(* IEC 61131-3 sources: RoboFlex-Cell/plc/codesys, 6 files *)

(* ---- FB_Alarm.st ---- *)
FUNCTION_BLOCK FB_Alarm
VAR_INPUT
    Trip : BOOL;
    Code : UINT;
    ResetAccepted : BOOL;
END_VAR
VAR_OUTPUT
    Active : BOOL;
    LatchedCode : UINT;
END_VAR
IF Trip THEN
    IF NOT Active THEN
        LatchedCode := Code;
    END_IF;
    Active := TRUE;
ELSIF ResetAccepted THEN
    Active := FALSE;
    LatchedCode := 0;
END_IF;
END_FUNCTION_BLOCK

(* ---- FB_Conveyor.st ---- *)
FUNCTION_BLOCK FB_Conveyor
VAR_INPUT
    RunRequest : BOOL;
    SafeEnable : BOOL;
    JamDetected : BOOL;
END_VAR
VAR_OUTPUT
    MotorRun : BOOL;
END_VAR
MotorRun := RunRequest AND SafeEnable AND NOT JamDetected;
END_FUNCTION_BLOCK

(* ---- FB_Gripper.st ---- *)
FUNCTION_BLOCK FB_Gripper
VAR_INPUT
    CloseRequest : BOOL;
    ClosedFeedback : BOOL;
    OpenFeedback : BOOL;
    SafeEnable : BOOL;
    Reset : BOOL;
END_VAR
VAR_OUTPUT
    CloseValve : BOOL;
    AtPosition : BOOL;
    Error : BOOL;
END_VAR
VAR
    FeedbackTimer : TON;
END_VAR
(* Hold the last valve command on a software safety stop; never drop a part.
   A physical safety circuit requires an independently assessed pneumatic design. *)
IF SafeEnable THEN
    CloseValve := CloseRequest;
END_IF;
AtPosition := (CloseRequest AND ClosedFeedback) OR (NOT CloseRequest AND OpenFeedback);
FeedbackTimer(IN := SafeEnable AND NOT AtPosition, PT := T#500ms);
IF Reset THEN
    Error := FALSE;
ELSIF FeedbackTimer.Q THEN
    Error := TRUE;
END_IF;
END_FUNCTION_BLOCK

(* ---- FB_Robot.st ---- *)
FUNCTION_BLOCK FB_Robot
VAR_INPUT
    Execute : BOOL;
    SafeEnable : BOOL;
    Reset : BOOL;
    Ready : BOOL;
    Running : BOOL;
    Complete : BOOL;
    RobotError : BOOL;
END_VAR
VAR_OUTPUT
    Start : BOOL;
    Ack : BOOL;
    Stop : BOOL;
    Done : BOOL;
    Error : BOOL;
    ErrorId : UINT;
END_VAR
VAR
    Phase : UINT;
    StartEdge : R_TRIG;
    StartTimer : TON;
    MotionTimer : TON;
    AckTimer : TON;
END_VAR

StartEdge(CLK := Execute);
StartTimer(IN := Phase = 10, PT := T#500ms);
MotionTimer(IN := Phase = 20, PT := T#6s);
AckTimer(IN := Phase = 30, PT := T#500ms);
Start := FALSE;
Ack := FALSE;
Stop := NOT SafeEnable;

IF Reset AND SafeEnable THEN
    Phase := 0;
    Done := FALSE;
    Error := FALSE;
    ErrorId := 0;
ELSIF NOT SafeEnable THEN
    Phase := 0;
    Done := FALSE;
ELSIF RobotError THEN
    Error := TRUE;
    ErrorId := 3;
END_IF;

IF SafeEnable AND NOT Reset AND NOT Error THEN
    CASE Phase OF
        0:
            IF StartEdge.Q THEN
                IF Ready AND NOT Complete AND NOT Running THEN
                    Phase := 10;
                ELSE
                    Error := TRUE;
                    ErrorId := 3;
                END_IF;
            END_IF;
        10:
            Start := TRUE;
            IF Running THEN
                Start := FALSE;
                Phase := 20;
            ELSIF StartTimer.Q THEN
                Error := TRUE;
                ErrorId := 4;
            END_IF;
        20:
            IF Complete AND NOT Running THEN
                Phase := 30;
            ELSIF MotionTimer.Q THEN
                Error := TRUE;
                ErrorId := 4;
            END_IF;
        30:
            Ack := TRUE;
            IF NOT Complete AND Ready THEN
                Ack := FALSE;
                Done := TRUE;
                Phase := 40;
            ELSIF AckTimer.Q THEN
                Error := TRUE;
                ErrorId := 4;
            END_IF;
        40:
            IF NOT Execute THEN
                Done := FALSE;
                Phase := 0;
            END_IF;
    END_CASE;
END_IF;
IF Error THEN
    Start := FALSE;
    Ack := FALSE;
    Stop := TRUE;
END_IF;
END_FUNCTION_BLOCK

(* ---- FB_Sequence.st ---- *)
FUNCTION_BLOCK FB_Sequence
VAR_INPUT
    StartButton : BOOL;
    StopButton : BOOL;
    ResetButton : BOOL;
    ManualPartClear : BOOL;
    SafetyOK : BOOL;
    HeartbeatOK : BOOL;
    PartDetected : BOOL;
    JamDetected : BOOL;
    VisionDone : BOOL;
    VisionError : BOOL;
    VisionErrorId : UINT;
    RobotDone : BOOL;
    RobotError : BOOL;
    RobotErrorId : UINT;
    GripperClosed : BOOL;
    GripperOpen : BOOL;
    GripperError : BOOL;
    QualityOK : BOOL;
END_VAR
VAR_OUTPUT
    State : UINT; (* 0 idle, 30 wait, 40 vision, 50 pick, 55 grip, 60 place,
                     65 release, 70 check, 75 home, 80 complete, 900 error *)
    ConveyorRequest : BOOL;
    VisionExecute : BOOL;
    RobotExecute : BOOL;
    JobNumber : UINT; (* 1 pick, 2 place, 3 home; pose data sent separately *)
    CloseRequest : BOOL;
    AlarmCode : UINT;
    ResetAccepted : BOOL;
    OKCount : UDINT;
    NGCount : UDINT;
END_VAR
VAR
    StartEdge : R_TRIG;
    ResetEdge : R_TRIG;
    StateTimer : TON;
    LastState : UINT;
    TripCode : UINT;
END_VAR

StartEdge(CLK := StartButton);
ResetEdge(CLK := ResetButton);
StateTimer(IN := State = LastState AND State <> 0 AND State <> 900, PT := T#2s);
LastState := State;
ResetAccepted := FALSE;
TripCode := 0;
ConveyorRequest := FALSE;
VisionExecute := FALSE;
RobotExecute := FALSE;

IF NOT SafetyOK THEN
    TripCode := 10; (* actual E-stop/door distinction belongs in mapped safety status *)
ELSIF State <> 0 AND State <> 900 THEN
    IF NOT HeartbeatOK THEN TripCode := 7;
    ELSIF StopButton THEN TripCode := 13;
    ELSIF RobotError THEN TripCode := RobotErrorId;
    ELSIF VisionError THEN TripCode := VisionErrorId;
    ELSIF GripperError THEN TripCode := 5;
    ELSIF JamDetected THEN TripCode := 9;
    END_IF;
END_IF;

IF TripCode <> 0 AND State <> 900 THEN
    AlarmCode := TripCode;
    State := 900;
END_IF;

CASE State OF
    0:
        IF StartEdge.Q AND SafetyOK AND HeartbeatOK AND NOT JamDetected THEN State := 30; END_IF;
    30:
        ConveyorRequest := TRUE;
        IF PartDetected THEN
            ConveyorRequest := FALSE;
            State := 40;
        ELSIF StateTimer.Q THEN
            AlarmCode := 8;
            State := 900;
        END_IF;
    40:
        VisionExecute := TRUE;
        IF VisionDone THEN State := 50; END_IF;
    50:
        JobNumber := 1;
        RobotExecute := TRUE;
        IF RobotDone THEN State := 55; END_IF;
    55:
        CloseRequest := TRUE;
        IF GripperClosed THEN State := 60; END_IF;
    60:
        JobNumber := 2;
        RobotExecute := TRUE;
        IF RobotDone THEN State := 65; END_IF;
    65:
        CloseRequest := FALSE;
        IF GripperOpen THEN State := 70; END_IF;
    70:
        IF QualityOK THEN State := 75;
        ELSIF StateTimer.Q THEN
            NGCount := NGCount + 1;
            AlarmCode := 6;
            State := 900;
        END_IF;
    75:
        JobNumber := 3;
        RobotExecute := TRUE;
        IF RobotDone THEN State := 80; END_IF;
    80:
        OKCount := OKCount + 1;
        State := 30;
    900:
        IF ResetEdge.Q AND SafetyOK AND HeartbeatOK AND NOT JamDetected AND ManualPartClear THEN
            ResetAccepted := TRUE;
            CloseRequest := FALSE;
            AlarmCode := 0;
            State := 0;
        END_IF;
END_CASE;
IF State = 900 THEN
    ConveyorRequest := FALSE;
    VisionExecute := FALSE;
    RobotExecute := FALSE;
END_IF;
END_FUNCTION_BLOCK

(* ---- FB_Vision.st ---- *)
FUNCTION_BLOCK FB_Vision
VAR_INPUT
    Execute : BOOL;
    SafeEnable : BOOL;
    Connected : BOOL;
    ResultValid : BOOL;
    ResultOK : BOOL;
    Reset : BOOL;
END_VAR
VAR_OUTPUT
    Trigger : BOOL;
    Ack : BOOL;
    Done : BOOL;
    Error : BOOL;
    ErrorId : UINT;
END_VAR
VAR
    Phase : UINT;
    Edge : R_TRIG;
    ResultTimer : TON;
    ClearTimer : TON;
END_VAR
Edge(CLK := Execute);
ResultTimer(IN := Phase = 10, PT := T#1s);
ClearTimer(IN := Phase = 20, PT := T#500ms);
Trigger := FALSE;
Ack := FALSE;
IF Reset OR NOT SafeEnable THEN
    Phase := 0;
    Done := FALSE;
    Error := FALSE;
    ErrorId := 0;
ELSIF NOT Error THEN
    CASE Phase OF
        0:
            IF Edge.Q THEN
                IF Connected AND NOT ResultValid THEN
                    Phase := 10;
                ELSE
                    Error := TRUE;
                    ErrorId := 1;
                END_IF;
            END_IF;
        10:
            Trigger := TRUE;
            IF NOT Connected THEN
                Error := TRUE;
                ErrorId := 1;
            ELSIF ResultValid THEN
                Trigger := FALSE;
                IF ResultOK THEN
                    Phase := 20;
                ELSE
                    Error := TRUE;
                    ErrorId := 2;
                END_IF;
            ELSIF ResultTimer.Q THEN
                Error := TRUE;
                ErrorId := 2;
            END_IF;
        20:
            Ack := TRUE;
            IF NOT ResultValid THEN
                Ack := FALSE;
                Done := TRUE;
                Phase := 30;
            ELSIF ClearTimer.Q THEN
                Error := TRUE;
                ErrorId := 2;
            END_IF;
        30:
            IF NOT Execute THEN
                Done := FALSE;
                Phase := 0;
            END_IF;
    END_CASE;
END_IF;
IF Error THEN
    Trigger := FALSE;
    Ack := FALSE;
END_IF;
END_FUNCTION_BLOCK
